TYPE ST_TriggerTellControl :
STRUCT
	sim	  	: BOOL;
	start 	: BOOL;
	reset	: BOOL;
END_STRUCT
END_TYPE

(* stored: Version 1.1.0.1, ProductVersion 3.1.4024.12
   DUT ST_TriggerTellControl: Id {35e2e531-dbc6-432d-a9cc-2c6cb9a29552} *)
